FUNCTION F_DecodeDriveState : E_DriveState
VAR_INPUT
    statusWord : UINT; // 0x6041
END_VAR
VAR
    masked : UINT;
END_VAR

masked := statusWord AND 16#006F;

IF (masked AND 16#0008) <> 0 THEN
    // bit3 = Fault
    F_DecodeDriveState := E_DriveState.FAULT;
ELSIF masked = 16#0060 THEN
    // Switch on disabled
    F_DecodeDriveState := E_DriveState.SWITCH_ON_DISABLED;
ELSIF masked = 16#0021 THEN
    // Ready to switch on
    F_DecodeDriveState := E_DriveState.READY_TO_SWITCH_ON;
ELSIF masked = 16#0023 THEN
    // Switched on
    F_DecodeDriveState := E_DriveState.SWITCHED_ON;
ELSIF masked = 16#0027 THEN
    // Operation enabled
    F_DecodeDriveState := E_DriveState.OPERATION_ENABLED;
ELSE
    F_DecodeDriveState := E_DriveState.UNKNOWN;
END_IF

END_FUNCTION

(* stored: Version 1.1.0.1
   POU F_DecodeDriveState: Id {c439a05c-b7ee-4ef5-8b86-661d59fe3393}, SpecialFunc None *)
